FUNCTION_BLOCK "Prova"
TITLE =
VERSION : 0.1

VAR_INPUT
  Avvio : Bool;
END_VAR

BEGIN
NETWORK
TITLE =
    FOO %I0.0;
	XX %I0.1;
	A %I0.2;
END_FUNCTION_BLOCK
